// TIA Portal V15.1 export
FUNCTION "HmiMap" : Void   // FC3, LAD
TITLE = HmiMap
{ S7_Optimized_Access := 'TRUE' }
VERSION : 0.1
// 0007 / H-05: alarm display map only; writes HmiAlm only, no Ack
// stored: AutoNumber false, IsIECCheckEnabled false, SetENOAutomatically False
BEGIN

REGION Network 1: C01 / 0007 H-05 — Common.x0: E-STOP active or not reset; clears: Release E-STOP and RESET
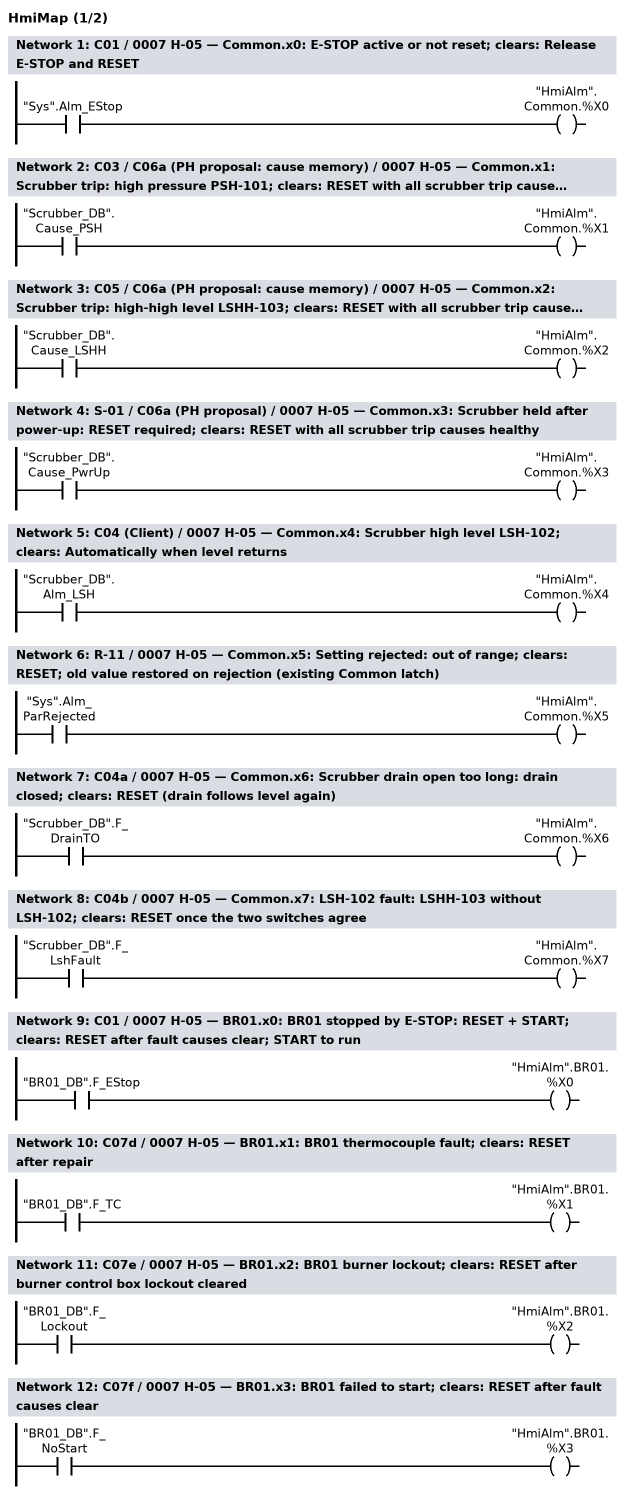
   RUNG wire#powerrail
      Contact( "Sys".Alm_EStop )
      Coil( "HmiAlm".Common.%X0 )
   END_RUNG
   // the same network as SCL:
   "HmiAlm".Common.%X0 := "Sys".Alm_EStop;
END_REGION

REGION Network 2: C03 / C06a (PH proposal: cause memory) / 0007 H-05 — Common.x1: Scrubber trip: high pressure PSH-101; clears: RESET with all scrubber trip causes healthy
   RUNG wire#powerrail
      Contact( "Scrubber_DB".Cause_PSH )
      Coil( "HmiAlm".Common.%X1 )
   END_RUNG
   // the same network as SCL:
   "HmiAlm".Common.%X1 := "Scrubber_DB".Cause_PSH;
END_REGION

REGION Network 3: C05 / C06a (PH proposal: cause memory) / 0007 H-05 — Common.x2: Scrubber trip: high-high level LSHH-103; clears: RESET with all scrubber trip causes healthy
   RUNG wire#powerrail
      Contact( "Scrubber_DB".Cause_LSHH )
      Coil( "HmiAlm".Common.%X2 )
   END_RUNG
   // the same network as SCL:
   "HmiAlm".Common.%X2 := "Scrubber_DB".Cause_LSHH;
END_REGION

REGION Network 4: S-01 / C06a (PH proposal) / 0007 H-05 — Common.x3: Scrubber held after power-up: RESET required; clears: RESET with all scrubber trip causes healthy
   RUNG wire#powerrail
      Contact( "Scrubber_DB".Cause_PwrUp )
      Coil( "HmiAlm".Common.%X3 )
   END_RUNG
   // the same network as SCL:
   "HmiAlm".Common.%X3 := "Scrubber_DB".Cause_PwrUp;
END_REGION

REGION Network 5: C04 (Client) / 0007 H-05 — Common.x4: Scrubber high level LSH-102; clears: Automatically when level returns
   RUNG wire#powerrail
      Contact( "Scrubber_DB".Alm_LSH )
      Coil( "HmiAlm".Common.%X4 )
   END_RUNG
   // the same network as SCL:
   "HmiAlm".Common.%X4 := "Scrubber_DB".Alm_LSH;
END_REGION

REGION Network 6: R-11 / 0007 H-05 — Common.x5: Setting rejected: out of range; clears: RESET; old value restored on rejection (existing Common latch)
   RUNG wire#powerrail
      Contact( "Sys".Alm_ParRejected )
      Coil( "HmiAlm".Common.%X5 )
   END_RUNG
   // the same network as SCL:
   "HmiAlm".Common.%X5 := "Sys".Alm_ParRejected;
END_REGION

REGION Network 7: C04a / 0007 H-05 — Common.x6: Scrubber drain open too long: drain closed; clears: RESET (drain follows level again)
   RUNG wire#powerrail
      Contact( "Scrubber_DB".F_DrainTO )
      Coil( "HmiAlm".Common.%X6 )
   END_RUNG
   // the same network as SCL:
   "HmiAlm".Common.%X6 := "Scrubber_DB".F_DrainTO;
END_REGION

REGION Network 8: C04b / 0007 H-05 — Common.x7: LSH-102 fault: LSHH-103 without LSH-102; clears: RESET once the two switches agree
   RUNG wire#powerrail
      Contact( "Scrubber_DB".F_LshFault )
      Coil( "HmiAlm".Common.%X7 )
   END_RUNG
   // the same network as SCL:
   "HmiAlm".Common.%X7 := "Scrubber_DB".F_LshFault;
END_REGION

REGION Network 9: C01 / 0007 H-05 — BR01.x0: BR01 stopped by E-STOP: RESET + START; clears: RESET after fault causes clear; START to run
   RUNG wire#powerrail
      Contact( "BR01_DB".F_EStop )
      Coil( "HmiAlm".BR01.%X0 )
   END_RUNG
   // the same network as SCL:
   "HmiAlm".BR01.%X0 := "BR01_DB".F_EStop;
END_REGION

REGION Network 10: C07d / 0007 H-05 — BR01.x1: BR01 thermocouple fault; clears: RESET after repair
   RUNG wire#powerrail
      Contact( "BR01_DB".F_TC )
      Coil( "HmiAlm".BR01.%X1 )
   END_RUNG
   // the same network as SCL:
   "HmiAlm".BR01.%X1 := "BR01_DB".F_TC;
END_REGION

REGION Network 11: C07e / 0007 H-05 — BR01.x2: BR01 burner lockout; clears: RESET after burner control box lockout cleared
   RUNG wire#powerrail
      Contact( "BR01_DB".F_Lockout )
      Coil( "HmiAlm".BR01.%X2 )
   END_RUNG
   // the same network as SCL:
   "HmiAlm".BR01.%X2 := "BR01_DB".F_Lockout;
END_REGION

REGION Network 12: C07f / 0007 H-05 — BR01.x3: BR01 failed to start; clears: RESET after fault causes clear
   RUNG wire#powerrail
      Contact( "BR01_DB".F_NoStart )
      Coil( "HmiAlm".BR01.%X3 )
   END_RUNG
   // the same network as SCL:
   "HmiAlm".BR01.%X3 := "BR01_DB".F_NoStart;
END_REGION

REGION Network 13: C07g / 0007 H-05 — BR01.x4: BR01 stopped by itself; clears: RESET after fault causes clear
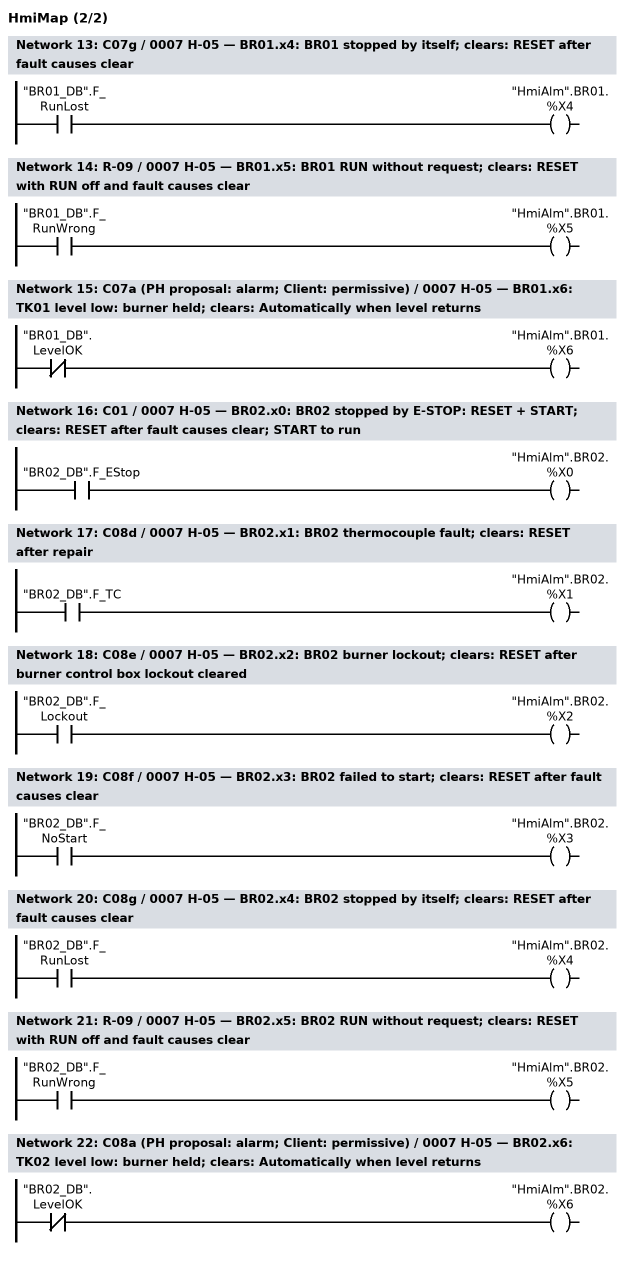
   RUNG wire#powerrail
      Contact( "BR01_DB".F_RunLost )
      Coil( "HmiAlm".BR01.%X4 )
   END_RUNG
   // the same network as SCL:
   "HmiAlm".BR01.%X4 := "BR01_DB".F_RunLost;
END_REGION

REGION Network 14: R-09 / 0007 H-05 — BR01.x5: BR01 RUN without request; clears: RESET with RUN off and fault causes clear
   RUNG wire#powerrail
      Contact( "BR01_DB".F_RunWrong )
      Coil( "HmiAlm".BR01.%X5 )
   END_RUNG
   // the same network as SCL:
   "HmiAlm".BR01.%X5 := "BR01_DB".F_RunWrong;
END_REGION

REGION Network 15: C07a (PH proposal: alarm; Client: permissive) / 0007 H-05 — BR01.x6: TK01 level low: burner held; clears: Automatically when level returns
   RUNG wire#powerrail
      I_Contact( "BR01_DB".LevelOK )
      Coil( "HmiAlm".BR01.%X6 )
   END_RUNG
   // the same network as SCL:
   "HmiAlm".BR01.%X6 := NOT "BR01_DB".LevelOK;
END_REGION

REGION Network 16: C01 / 0007 H-05 — BR02.x0: BR02 stopped by E-STOP: RESET + START; clears: RESET after fault causes clear; START to run
   RUNG wire#powerrail
      Contact( "BR02_DB".F_EStop )
      Coil( "HmiAlm".BR02.%X0 )
   END_RUNG
   // the same network as SCL:
   "HmiAlm".BR02.%X0 := "BR02_DB".F_EStop;
END_REGION

REGION Network 17: C08d / 0007 H-05 — BR02.x1: BR02 thermocouple fault; clears: RESET after repair
   RUNG wire#powerrail
      Contact( "BR02_DB".F_TC )
      Coil( "HmiAlm".BR02.%X1 )
   END_RUNG
   // the same network as SCL:
   "HmiAlm".BR02.%X1 := "BR02_DB".F_TC;
END_REGION

REGION Network 18: C08e / 0007 H-05 — BR02.x2: BR02 burner lockout; clears: RESET after burner control box lockout cleared
   RUNG wire#powerrail
      Contact( "BR02_DB".F_Lockout )
      Coil( "HmiAlm".BR02.%X2 )
   END_RUNG
   // the same network as SCL:
   "HmiAlm".BR02.%X2 := "BR02_DB".F_Lockout;
END_REGION

REGION Network 19: C08f / 0007 H-05 — BR02.x3: BR02 failed to start; clears: RESET after fault causes clear
   RUNG wire#powerrail
      Contact( "BR02_DB".F_NoStart )
      Coil( "HmiAlm".BR02.%X3 )
   END_RUNG
   // the same network as SCL:
   "HmiAlm".BR02.%X3 := "BR02_DB".F_NoStart;
END_REGION

REGION Network 20: C08g / 0007 H-05 — BR02.x4: BR02 stopped by itself; clears: RESET after fault causes clear
   RUNG wire#powerrail
      Contact( "BR02_DB".F_RunLost )
      Coil( "HmiAlm".BR02.%X4 )
   END_RUNG
   // the same network as SCL:
   "HmiAlm".BR02.%X4 := "BR02_DB".F_RunLost;
END_REGION

REGION Network 21: R-09 / 0007 H-05 — BR02.x5: BR02 RUN without request; clears: RESET with RUN off and fault causes clear
   RUNG wire#powerrail
      Contact( "BR02_DB".F_RunWrong )
      Coil( "HmiAlm".BR02.%X5 )
   END_RUNG
   // the same network as SCL:
   "HmiAlm".BR02.%X5 := "BR02_DB".F_RunWrong;
END_REGION

REGION Network 22: C08a (PH proposal: alarm; Client: permissive) / 0007 H-05 — BR02.x6: TK02 level low: burner held; clears: Automatically when level returns
   RUNG wire#powerrail
      I_Contact( "BR02_DB".LevelOK )
      Coil( "HmiAlm".BR02.%X6 )
   END_RUNG
   // the same network as SCL:
   "HmiAlm".BR02.%X6 := NOT "BR02_DB".LevelOK;
END_REGION
END_FUNCTION
